PROGRAM PRG_Tests
VAR
    fbLightTests : FB_LightTests;
	fbButtonTests : FB_ButtonTests;
    fbWorkshopTests : FB_WorkshopTests;
    fbHomeTests : FB_HomeTests;
    fbLightCatalogTests : FB_LightCatalogTests;
    fbLocalIntegrationTests : FB_LocalIntegrationTests;
    fbLightCommandTests : FB_LightCommandTests;
    fbMqttLightProtocolTests : FB_MqttLightProtocolTests;
    fbMqttConfigParserTests : FB_MqttConfigParserTests;
    fbMqttIntegrationQueueTests : FB_MqttIntegrationQueueTests;
    fbMqttDiscoveryTests : FB_MqttDiscoveryTests;
END_VAR

TcUnit.RUN();

END_PROGRAM

(* stored: Version 1.1.0.1
   POU PRG_Tests: Id {C914D478-7D86-472A-8A10-7D6FD9048733}, SpecialFunc None *)
